// SPS -> GUI. Status eines Niederhalters.
{attribute 'pack_mode' := '1'}
TYPE ST_HmiClampStatus :
STRUCT
    eState : E_ClampState;
    bValve : BOOL; // Ausgang
    bOpen : BOOL; // Endlage OFFEN
    fLastSwitchTime_ms : LREAL;
END_STRUCT
END_TYPE

(* stored: Version 1.1.0.1
   DUT ST_HmiClampStatus: Id {46c853e3-1ef2-4445-b91d-047126fb6a74} *)
